(* PLC project Motor_Control, PLCAutoPilot Machine Expert Logic Builder V19.2.3.0, author PLCAutoPilot *)
(* stored: creationDateTime 2025-12-30T03:00:00.0000000, version 1.0.0.0, modificationDateTime 2025-12-30T03:00:00.0000000 *)

PROGRAM Motor_Control_LD
  VAR
    StartPB AT %IX0.0 : BOOL;
    StopPB AT %IX0.1 : BOOL;
    MotorOut AT %QX0.0 : BOOL;
  END_VAR
  VAR
    StartupTimer : TON;
  END_VAR

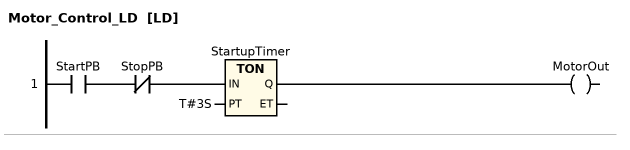
(* LD diagram, written out as Structured Text *)

StartupTimer(IN := StartPB AND NOT StopPB, PT := T#3S);
MotorOut := StartupTimer.Q;
END_PROGRAM
